Fanuc KAREL source: KT00927.KL

PROGRAM KT00927
%NOLOCKGROUP
VAR
  H1: ARRAY[2] OF SHORT
  H2: ARRAY[2] OF SHORT
  OUT: STRING[80]
BEGIN
  H1[1] = 2
  H2[1] = 3
  H1[1] = 2
  H2[1] = 3
  OUT = SUB_STR(H1[1], 1, 1)
END KT00927
